SUBAPPLICATION VarInOutSubappInterface
  (* Standard: 61499-1; Description: Copyright (c) 2026 Martin Erich Jobst This program and the accompanying materials are made available under the terms of the Eclipse Public License 2.0 which is available at https://www.eclipse.org/legal/epl-2.0/ SPDX-License-Identifier: EPL-2.0 *)
  (* Version 1.0, 2026-11-18, Martin Jobst *)
  PACKAGE lib::VarDeclaration;
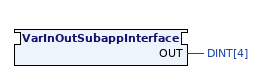
  VAR_OUTPUT
    OUT : ARRAY [0..3] OF DINT;
  END_VAR
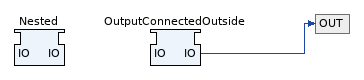
  SUBAPPLICATION Nested
    VAR_IN_OUT
      IO : ARRAY [0..3] OF DINT;
    END_VAR
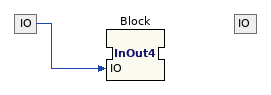
    FBS
      Block : lib::VarDeclaration::support::InOut4;
    END_FBS
    DATA_CONNECTIONS
      IO TO Block.IO;
    END_CONNECTIONS
  END_SUBAPPLICATION
  SUBAPPLICATION OutputConnectedOutside
    VAR_IN_OUT
      IO : ARRAY [0..3] OF DINT;
    END_VAR
  END_SUBAPPLICATION
  DATA_CONNECTIONS
    OutputConnectedOutside.IO TO OUT;
  END_CONNECTIONS
END_SUBAPPLICATION
